Fanuc KAREL source: KA00192.KL

PROGRAM KA00192
%NOLOCKGROUP
VAR
  SRC: ARRAY[4] OF SHORT
  DST: ARRAY[4] OF BOOLEAN
BEGIN
  DST = SRC
END KA00192
